(*
SPDX-FileCopyrightText: © 2026 Oleksandr Tiutyk <trofimich@gmail.com>
SPDX-License-Identifier: MIT
License: https://opensource.org/license/mit
*)

(*!
<summary>
Beckhoff 3-phase power measurement output control channel process image.
</summary>
<description>
One UINT8 Index selector at 0x7000:01, 0x7010:01 or 0x7020:01.
Common indices 0..5 select apparent power, reactive power, energy, power factor, frequency and negative energy.
Other indices depend on terminal/firmware. Wait for input acknowledgement and valid status before interpreting
VariantValue; a selector write is not a synchronous measurement read. Use one owner task for output writes.
When used for I/O, link located fields or their containing buffers to the matching selected PDOs.
The record is not a packed wire buffer; compiler padding is not part of the device specification.
Unlinked/default values do not prove valid I/O. The caller evaluates bus/channel validity before use.
Use one owner task per instance and externally synchronize other access; multi-field snapshots are not atomic.
Copies store data without creating hardware links. Keep borrowed field references valid while consumers are bound.
This passive record performs no validation, synchronization, configuration or protocol advancement.
</description>
*)
TYPE POWER_MEASUREMENT_OUTPUT_CHANNEL :
STRUCT
	Index AT %Q* : USINT;
END_STRUCT
END_TYPE

(* stored: Version 1.1.0.1, ProductVersion 3.1.4026.20
   DUT POWER_MEASUREMENT_OUTPUT_CHANNEL: Id {de115164-6cb4-496c-b03a-53db6a3d0569} *)
